TYPE Vector3 :
STRUCT
	x : LREAL;
	y : LREAL;
	z : LREAL;
END_STRUCT
END_TYPE

(* stored: Version 1.1.0.1, ProductVersion 3.1.4026.12
   DUT Vector3: Id {89307baf-b3c4-55e9-a3b9-13f2e3138d73} *)
